Fanuc KAREL source: kc00040.KL

-- PROVISIONAL review KL for V770-1; original PC SHA256 02b6b6d6b516e7dac10f3be222f507165f7248f840551e26b082339869af2305
-- Incomplete behavior may be omitted. Consult companion uncertainty JSON. Do not deploy.
PROGRAM KC00040
%NOLOCKGROUP
BEGIN
  -- UNRESOLVED_PC offsets 5-33; opcodes 27,22,22,22,22,31
  -- UNRESOLVED_PC offsets 38-42; opcodes 7F
END KC00040
